Staubli VAL3: bind_edit.pgx

program bind_edit()
  local num l_i
  local string l_sbtn
begin
  for l_i = 0 to size(bEditBool)-1
    l_sbtn="btn"+toString("",l_i)
    userPageBindClick("editProg",l_sbtn,bEditBool[l_i],true)
  endFor

  userPageBindClick("editProg","btnback",bEditBack,true)

  userPageBind("editProg","lbleditindex","innerHTML",sEditIndex,1,"r")
  userPageBind("editProg","lbleditpage","innerHTML",sEditPage,1,"r")

  userPageBind("editProg","lst1","value",sSelTRAJ,1,"rw")
end
